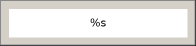
VISUALIZATION vis_IconState  // 196x46
VAR_IN_OUT
	value: INT;
END_VAR
VAR_INPUT
	reqValue: INT;
	text: STRING;	
END_VAR
    Rectangle (0,0 196x46), colour toggle: value=reqValue
    Textfield (8,8 180x30), "%s", text variable: text
        OnMouseClick: execute { value:=reqValue; }
END_VISUALIZATION

(* stored: Version 1.1.0.1, ProductVersion 3.1.4024.12
   Visu vis_IconState: Id {4dfee271-54cc-4dba-8d3d-68b6171f5d67} *)
